Universal Robots URScript: FeatureTest.script

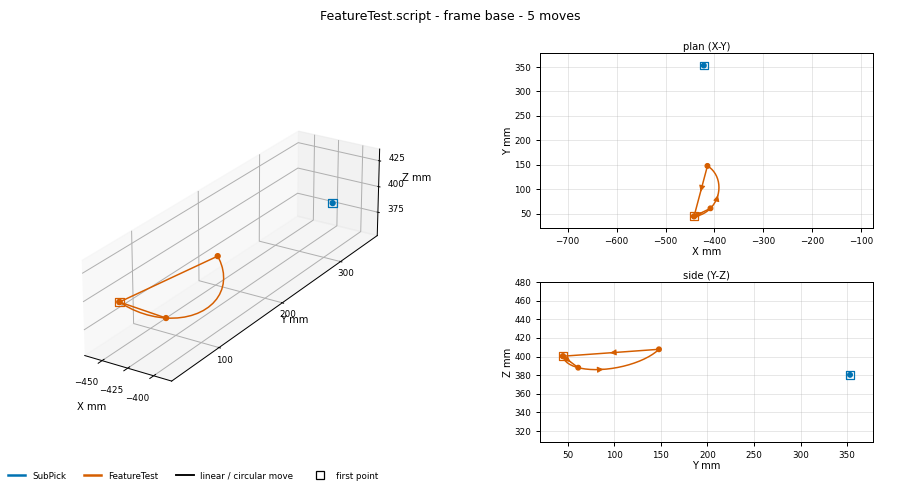
[picture p0: tool path of FeatureTest.script in frame base, 5 of 7 moves have a stored position in this frame; points joined in program order, loops and branches not executed]
def FeatureTest():
  # Global parameters:
  global speed_ms    = 0.250
  global speed_rads  = 0.750
  global accel_mss   = 1.200
  global accel_radss = 1.200
  global blend_radius_m = 0.001
  global ref_frame = p[0,0,0,0,0,0]

  #
  # TO REMOVE HEADER:
  # Go to "Program" -> "Post-Processor Editor"
  # Select "Universal Robots"
  # Set "INCLUDE_HEADER" to "False"
  #
  #--------------------------
  # Add any default subprograms here
  # For example, to drive a gripper as a program call:
  # def Gripper_Open():
  #   ...
  # end
  #
  # Example to drive a spray gun:
  def SprayOn(value):
    # use the value as an output:
    DO_SPRAY = 5
    if value == 0:
      set_standard_digital_out(DO_SPRAY, False)
    else:
      set_standard_digital_out(DO_SPRAY, True)
    end
  end

  # Example to drive an extruder:
  def Extruder(value):
    # use the value as an output:
    if value < 0:
      # stop extruder
    else:
      # start extruder
    end
  end

  # Example to move an external axis
  def MoveAxis(value):
    # use the value as an output:
    DO_AXIS_1 = 1
    DI_AXIS_1 = 1
    if value <= 0:
      set_standard_digital_out(DO_AXIS_1, False)

      # Wait for digital input to change state
      #while (get_standard_digital_in(DI_AXIS_1) != False):
      #  sync()
      #end
    else:
      set_standard_digital_out(DO_AXIS_1, True)

      # Wait for digital input to change state
      #while (get_standard_digital_in(DI_AXIS_1) != True):
      #  sync()
      #end
    end
  end
  #--------------------------

  # Subprogram SubPick
  def SubPick():
    movel(pose_trans(ref_frame,p[-0.421760, 0.353029, 0.380392, 3.048452, 0.496356, 0.454618]),accel_mss,speed_ms,0,0.000)
    set_standard_digital_out(7, True)
  end


  # Main program:
  # Program generated by VerticalBot Studio for UR5e on 25/10/2026 12:00:00
  # Using nominal kinematics.
  ref_frame = p[0.100000, -0.050000, 0.020000, 0.000000, 0.000000, 0.523599]
  set_tcp(p[0.010000, 0.000000, 0.120000, 0.000000, 0.261799, 0.000000])
  speed_ms    = 0.300
  speed_rads  = 1.571
  accel_mss   = 1.500
  accel_radss = 6.981
  blend_radius_m = 0.005
  movej([-0.523599, -1.745329, 1.570796, -1.396263, -1.570796, 0.349066],accel_radss,speed_rads,0,0.005)
  movel(pose_trans(ref_frame,p[-0.421760, 0.353029, 0.380392, 3.048452, 0.496356, 0.454618]),accel_mss,speed_ms,0,0.005)
  movec(pose_trans(ref_frame,p[-0.384494, 0.350433, 0.368074, 3.036811, 0.389569, 0.461666]),pose_trans(ref_frame,p[-0.346512, 0.428592, 0.387797, 3.069709, 0.117165, 0.434828]),accel_mss,speed_ms,0) # end trace
  speed_ms    = 0.050
  blend_radius_m = 0.000
  movel(pose_trans(ref_frame,p[-0.421760, 0.353029, 0.380392, 3.048452, 0.496356, 0.454618]),accel_mss,speed_ms,0,0.000)
  blend_radius_m = 0.000
  speed_ms    = 0.300
  movel(pose_trans(ref_frame,p[-0.384494, 0.350433, 0.368074, 3.036811, 0.389569, 0.461666]),accel_mss,speed_ms,0,0.000)
  set_standard_digital_out(3, True)
  DO_GRIP = 0
  while (get_standard_digital_in(5) != True):
    sync()
  end
  while (DI_PART != True):
    sync()
  end
  sleep(0.500)
  # a comment line
  popup("Hello operator","Message",False,False,blocking=False)
  MyFunc()
  SetRPM(5000)
  RAW_CODE_LINE
  SubPick()
  speed_rads  = 0.785
  set_tcp(p[0.010000, 0.000000, 0.120000, 0.000000, 0.261799, 0.000000])
  # Attach to Tool 1
  movej([-0.523599, -1.745329, 1.570796, -1.396263, -1.570796, 0.349066],accel_radss,speed_rads,0,0.000)
  halt() # reimplement this function to force stop
  # End of main program
end

FeatureTest()
